(* PLC project TBEN_L5_PLC11.project, CODESYS CODESYS V3.5 SP21 Patch 1 *)
(* stored: creationDateTime 2026-11-07T15:34:50.940518, modificationDateTime 2026-11-07T15:09:07.4034196 *)

{attribute 'qualified_only'}
// Bước handshake của client FB_IolCall
TYPE E_IolCallStep :
(
    IDLE := 0,
    WAIT := 1,    // đã vào hàng đợi master, chờ kết quả
    DONE := 2,
    ERR  := 3
) INT;
END_TYPE
